Fanuc KAREL source: kd00016.compact.KL

PROGRAM KD00016
%STACKSIZE=65535
%PRIORITY=65535
%NOLOCKGROUP
VAR
I : INTEGER
J : INTEGER
B : BOOLEAN
R : REAL
S : STRING[80]
BEGIN
I=0
CONNECT TIMER TO I
END KD00016
